FUNCTION_BLOCK IOTest16_HMI (* Service Interface Function Block Type *)
  (* Standard: 61499-2 *)
  (* Version 0.0, 11/13/2026, Sandeep Patil, Flexbridge AB, template *)
  PACKAGE Flexbridge.FestoMPS400;
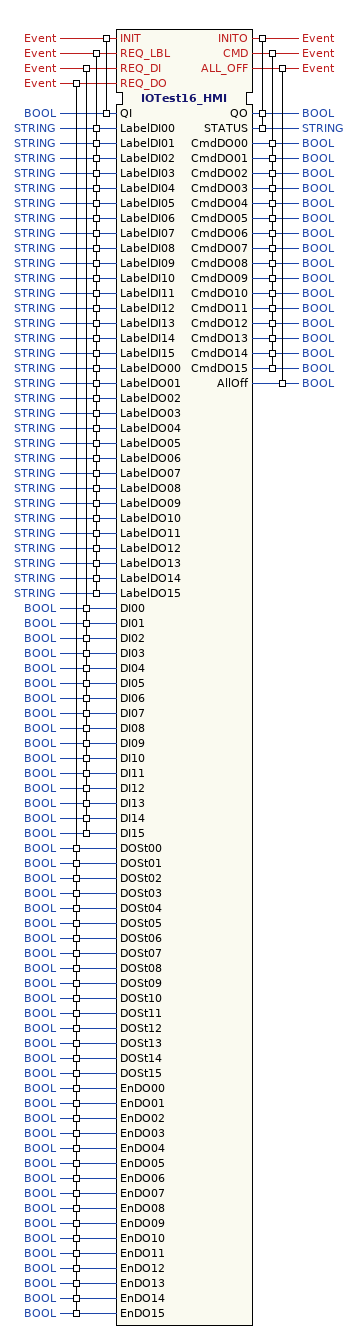
  EVENT_INPUT
    INIT WITH QI;
    REQ_LBL WITH LabelDI00, LabelDI01, LabelDI02, LabelDI03, LabelDI04, LabelDI05, LabelDI06, LabelDI07, LabelDI08, LabelDI09, LabelDI10, LabelDI11, LabelDI12, LabelDI13, LabelDI14, LabelDI15, LabelDO00, LabelDO01, LabelDO02, LabelDO03, LabelDO04, LabelDO05, LabelDO06, LabelDO07, LabelDO08, LabelDO09, LabelDO10, LabelDO11, LabelDO12, LabelDO13, LabelDO14, LabelDO15;
    REQ_DI WITH DI00, DI01, DI02, DI03, DI04, DI05, DI06, DI07, DI08, DI09, DI10, DI11, DI12, DI13, DI14, DI15;
    REQ_DO WITH DOSt00, DOSt01, DOSt02, DOSt03, DOSt04, DOSt05, DOSt06, DOSt07, DOSt08, DOSt09, DOSt10, DOSt11, DOSt12, DOSt13, DOSt14, DOSt15, EnDO00, EnDO01, EnDO02, EnDO03, EnDO04, EnDO05, EnDO06, EnDO07, EnDO08, EnDO09, EnDO10, EnDO11, EnDO12, EnDO13, EnDO14, EnDO15;
  END_EVENT
  EVENT_OUTPUT
    INITO WITH QO, STATUS;
    CMD WITH CmdDO00, CmdDO01, CmdDO02, CmdDO03, CmdDO04, CmdDO05, CmdDO06, CmdDO07, CmdDO08, CmdDO09, CmdDO10, CmdDO11, CmdDO12, CmdDO13, CmdDO14, CmdDO15;
    ALL_OFF WITH AllOff;
  END_EVENT
  VAR_INPUT
    QI : BOOL;
    LabelDI00 : STRING; (* Label text *)
    LabelDI01 : STRING; (* Label text *)
    LabelDI02 : STRING; (* Label text *)
    LabelDI03 : STRING; (* Label text *)
    LabelDI04 : STRING; (* Label text *)
    LabelDI05 : STRING; (* Label text *)
    LabelDI06 : STRING; (* Label text *)
    LabelDI07 : STRING; (* Label text *)
    LabelDI08 : STRING; (* Label text *)
    LabelDI09 : STRING; (* Label text *)
    LabelDI10 : STRING; (* Label text *)
    LabelDI11 : STRING; (* Label text *)
    LabelDI12 : STRING; (* Label text *)
    LabelDI13 : STRING; (* Label text *)
    LabelDI14 : STRING; (* Label text *)
    LabelDI15 : STRING; (* Label text *)
    LabelDO00 : STRING; (* Label text *)
    LabelDO01 : STRING; (* Label text *)
    LabelDO02 : STRING; (* Label text *)
    LabelDO03 : STRING; (* Label text *)
    LabelDO04 : STRING; (* Label text *)
    LabelDO05 : STRING; (* Label text *)
    LabelDO06 : STRING; (* Label text *)
    LabelDO07 : STRING; (* Label text *)
    LabelDO08 : STRING; (* Label text *)
    LabelDO09 : STRING; (* Label text *)
    LabelDO10 : STRING; (* Label text *)
    LabelDO11 : STRING; (* Label text *)
    LabelDO12 : STRING; (* Label text *)
    LabelDO13 : STRING; (* Label text *)
    LabelDO14 : STRING; (* Label text *)
    LabelDO15 : STRING; (* Label text *)
    DI00 : BOOL; (* Input lamp *)
    DI01 : BOOL; (* Input lamp *)
    DI02 : BOOL; (* Input lamp *)
    DI03 : BOOL; (* Input lamp *)
    DI04 : BOOL; (* Input lamp *)
    DI05 : BOOL; (* Input lamp *)
    DI06 : BOOL; (* Input lamp *)
    DI07 : BOOL; (* Input lamp *)
    DI08 : BOOL; (* Input lamp *)
    DI09 : BOOL; (* Input lamp *)
    DI10 : BOOL; (* Input lamp *)
    DI11 : BOOL; (* Input lamp *)
    DI12 : BOOL; (* Input lamp *)
    DI13 : BOOL; (* Input lamp *)
    DI14 : BOOL; (* Input lamp *)
    DI15 : BOOL; (* Input lamp *)
    DOSt00 : BOOL; (* Output state lamp *)
    DOSt01 : BOOL; (* Output state lamp *)
    DOSt02 : BOOL; (* Output state lamp *)
    DOSt03 : BOOL; (* Output state lamp *)
    DOSt04 : BOOL; (* Output state lamp *)
    DOSt05 : BOOL; (* Output state lamp *)
    DOSt06 : BOOL; (* Output state lamp *)
    DOSt07 : BOOL; (* Output state lamp *)
    DOSt08 : BOOL; (* Output state lamp *)
    DOSt09 : BOOL; (* Output state lamp *)
    DOSt10 : BOOL; (* Output state lamp *)
    DOSt11 : BOOL; (* Output state lamp *)
    DOSt12 : BOOL; (* Output state lamp *)
    DOSt13 : BOOL; (* Output state lamp *)
    DOSt14 : BOOL; (* Output state lamp *)
    DOSt15 : BOOL; (* Output state lamp *)
    EnDO00 : BOOL; (* Button enabled *)
    EnDO01 : BOOL; (* Button enabled *)
    EnDO02 : BOOL; (* Button enabled *)
    EnDO03 : BOOL; (* Button enabled *)
    EnDO04 : BOOL; (* Button enabled *)
    EnDO05 : BOOL; (* Button enabled *)
    EnDO06 : BOOL; (* Button enabled *)
    EnDO07 : BOOL; (* Button enabled *)
    EnDO08 : BOOL; (* Button enabled *)
    EnDO09 : BOOL; (* Button enabled *)
    EnDO10 : BOOL; (* Button enabled *)
    EnDO11 : BOOL; (* Button enabled *)
    EnDO12 : BOOL; (* Button enabled *)
    EnDO13 : BOOL; (* Button enabled *)
    EnDO14 : BOOL; (* Button enabled *)
    EnDO15 : BOOL; (* Button enabled *)
  END_VAR
  VAR_OUTPUT
    QO : BOOL; (* Event Output Qualifier *)
    STATUS : STRING; (* Service Status *)
    CmdDO00 : BOOL; (* Button: requested output state *)
    CmdDO01 : BOOL; (* Button: requested output state *)
    CmdDO02 : BOOL; (* Button: requested output state *)
    CmdDO03 : BOOL; (* Button: requested output state *)
    CmdDO04 : BOOL; (* Button: requested output state *)
    CmdDO05 : BOOL; (* Button: requested output state *)
    CmdDO06 : BOOL; (* Button: requested output state *)
    CmdDO07 : BOOL; (* Button: requested output state *)
    CmdDO08 : BOOL; (* Button: requested output state *)
    CmdDO09 : BOOL; (* Button: requested output state *)
    CmdDO10 : BOOL; (* Button: requested output state *)
    CmdDO11 : BOOL; (* Button: requested output state *)
    CmdDO12 : BOOL; (* Button: requested output state *)
    CmdDO13 : BOOL; (* Button: requested output state *)
    CmdDO14 : BOOL; (* Button: requested output state *)
    CmdDO15 : BOOL; (* Button: requested output state *)
    AllOff : BOOL; (* Button: all outputs off *)
  END_VAR
  SERVICE /
    SEQUENCE 
    END_SEQUENCE
  END_SERVICE
END_FUNCTION_BLOCK
